Fanuc KAREL source: KD00062.KL

PROGRAM KD00062
%NOLOCKGROUP
VAR
  I: INTEGER
  J: INTEGER
  B: BOOLEAN
  R: REAL
  S: STRING[80]
BEGIN
  CONDITION[1]:
  WHEN DIN[1] = ON DO
    ENABLE CONDITION[1]
  ENDCONDITION
END KD00062
